VISUALIZATION NavBar  // 1024x768
END_VISUALIZATION

(* stored: Version 1.1.0.1
   Visu NavBar: Id {5c55a31d-f689-43c4-bb2e-1c218b673ce8} *)
